VISUALIZATION CNV_Settings  // 1024x768
END_VISUALIZATION

(* stored: Version 1.1.0.1
   Visu CNV_Settings: Id {ec89c1b7-7a20-4c98-b2d4-743b830b709c} *)
